FUNCTION_BLOCK "Q08"
VERSION : 0.1
VAR_INPUT
    count : DINT;
END_VAR
VAR_IN_OUT
    analogValues : ARRAY[*] OF INT;
    channels : ARRAY[*] OF ST_AnalogChannel;
END_VAR
BEGIN
END_FUNCTION_BLOCK
